(* PLC project Vn_fanout_int, Beckhoff Automation GmbH TwinCAT PLC Control 3.5.13.21 *)
(* stored: creationDateTime 1970-01-01T00:00:00 *)

PROGRAM Vn_fanout_int
  VAR  (* added by the conversion: wires and edge detectors of the diagram *)
    _ADD10000000003_OUT : ANY;
  END_VAR

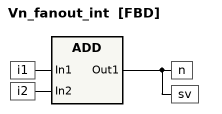
(* FBD diagram, written out as Structured Text *)
_ADD10000000003_OUT := i1 + i2;
n := _ADD10000000003_OUT;
sv := _ADD10000000003_OUT;
END_PROGRAM
